# B&R Automation Studio project 67
Automation Studio 4.12.10.39

## Configuration Config1

CPU 4PP065.0571-P74, AutomationRuntime D4.52, Build 4.1.2, Vc V4.52.0

### Task classes (Cpu.sw)
```
Cyclic#1:
  Program <- Program.prg
Libraries: Library
```

### Hardware
```
4PP065_0571_P74 : 4PP065.0571-P74 v1.2.0.0
  Connector IF4:
    DNAConfiguration = manual
  Connector IF5:
    ActivateDevice = 1
  ConfigurationID = 67_Config1
  Simulation = 1
  SystemTick = 10000
  TaskClassIdleTime = 10000
```

- Physical/Config1/4PP065_0571_P74/IoMap.iom: same as Physical/Config1/4PP065_0571_P74/Cpu.per
- Physical/Config1/4PP065_0571_P74/PvMap.vvm: same as Physical/Config1/4PP065_0571_P74/Cpu.per
## Logical view

Binary libraries used (declarations not repeated): operator, runtime, astime, AsIecCon


### Program Logical/Program (ANSIC)

#### main.c - Cyclic code
```c
#include <bur/plctypes.h>

#ifdef _DEFAULT_INCLUDES
	#include <AsDefault.h>
#endif

void _CYCLIC ProgramCyclic(void)
{
	counter++;
	if (counter >= 1100)
	{
		counter = 0;
	}

	if ((counter >= 100)&&(counter < 600))
	{
		Speed = 100.0;
	}
	else
	{
		Speed = 0.0;
	}

	if (Enable)
	{
		fb_controller.e = Speed - fb_motor.w;
		FB_Regulator(&fb_controller);

		fb_motor.u = fb_controller.u;
		FB_Motor(&fb_motor);

		fb_motor2.u = Speed * fb_motor2.ke;
		FB_Motor(&fb_motor2);
	}
}
```

#### Init.c - Initialization code
```c
#include <bur/plctypes.h>

#ifdef _DEFAULT_INCLUDES
	#include <AsDefault.h>
#endif

void _INIT ProgramInit(void)
{
	//LEGO NXT

	fb_motor.tm = 0.081;
	fb_motor.ke = 0.0641;
	fb_motor.dt = 0.01;

	fb_motor.w = 0.0;
	fb_motor.phi = 0.0;
	fb_motor.integrator.in = 0.0;
	fb_motor.integrator.out = 0.0;
	fb_motor.integrator.dt = 0.01;

	fb_motor2.tm = 0.081;
	fb_motor2.ke = 0.0641;
	fb_motor2.dt = 0.01;

	fb_motor2.w = 0.0;
	fb_motor2.phi = 0.0;
	fb_motor2.integrator.in = 0.0;
	fb_motor2.integrator.out = 0.0;
	fb_motor2.integrator.dt = 0.01;

	fb_controller.k_p = 0.0052;	/* ke*Tm/Tj, Tj = 1 s */
	fb_controller.k_i = 0.0641;	/* ke/Tj */
	fb_controller.max_abs_value = 9.0;
	fb_controller.dt = 0.01;

	fb_controller.iyOld = 0.0;
	fb_controller.integrator.in = 0.0;
	fb_controller.integrator.out = 0.0;
	fb_controller.integrator.dt = 0.01;

	Speed = 0.0;
	Enable = 1;
	counter = 0;

}
```

#### Exit.c - Exit code
```c
#include <bur/plctypes.h>

#ifdef _DEFAULT_INCLUDES
	#include <AsDefault.h>
#endif

void _EXIT ProgramExit(void)
{

}
```

#### Variables.var - Local variables
```iecst
VAR
	fb_controller : {REDUND_UNREPLICABLE} FB_Regulator;
	fb_motor : {REDUND_UNREPLICABLE} FB_Motor;
	Speed : {REDUND_UNREPLICABLE} REAL;
	Enable : {REDUND_UNREPLICABLE} BOOL;
	fb_motor2 : {REDUND_UNREPLICABLE} FB_Motor;
	counter : {REDUND_UNREPLICABLE} UDINT;
END_VAR
```

### Library Logical/Library (ANSIC)

#### Library.fun - Exported functions and function blocks
```iecst
{REDUND_ERROR} {REDUND_UNREPLICABLE} FUNCTION_BLOCK FB_Integrator (*Интегратор*) (*$GROUP=User,$CAT=User,$GROUPICON=User.png,$CATICON=User.png*)
	VAR_INPUT
		in : {REDUND_UNREPLICABLE} REAL; (*Вход интегратора*)
	END_VAR
	VAR_OUTPUT
		out : {REDUND_UNREPLICABLE} REAL; (*Выход интегратора*)
	END_VAR
	VAR
		dt : {REDUND_UNREPLICABLE} REAL; (*Шаг расчёта, с*)
	END_VAR
END_FUNCTION_BLOCK

{REDUND_ERROR} {REDUND_UNREPLICABLE} FUNCTION_BLOCK FB_Motor (*Модель ДПТ*) (*$GROUP=User,$CAT=User,$GROUPICON=User.png,$CATICON=User.png*)
	VAR_INPUT
		u : {REDUND_UNREPLICABLE} REAL; (*Напряжение, В*)
	END_VAR
	VAR_OUTPUT
		w : {REDUND_UNREPLICABLE} REAL; (*Частота вращения, об/мин*)
		phi : {REDUND_UNREPLICABLE} REAL; (*Положение вала*)
	END_VAR
	VAR
		integrator : {REDUND_UNREPLICABLE} FB_Integrator; (*Интегратор*)
		tm : {REDUND_UNREPLICABLE} REAL; (*Электромеханическая постоянная времени, с*)
		ke : {REDUND_UNREPLICABLE} REAL; (*Постоянная ЭДС, В*мин/об*)
		dt : {REDUND_UNREPLICABLE} REAL; (*Шаг расчёта, с*)
	END_VAR
END_FUNCTION_BLOCK

{REDUND_ERROR} {REDUND_UNREPLICABLE} FUNCTION_BLOCK FB_Regulator (*ПИ-регулятор*) (*$GROUP=User,$CAT=User,$GROUPICON=User.png,$CATICON=User.png*)
	VAR_INPUT
		e : {REDUND_UNREPLICABLE} REAL; (*Ошибка, об/мин*)
	END_VAR
	VAR_OUTPUT
		u : {REDUND_UNREPLICABLE} REAL; (*Напряжение на ДПТ, В*)
	END_VAR
	VAR
		k_p : {REDUND_UNREPLICABLE} REAL; (*Пропорциональный коэффициент*)
		k_i : {REDUND_UNREPLICABLE} REAL; (*Интегральный коэффициент*)
		integrator : {REDUND_UNREPLICABLE} FB_Integrator; (*Интегратор*)
		iyOld : {REDUND_UNREPLICABLE} REAL; (*Интегральная составляющая*)
		max_abs_value : {REDUND_UNREPLICABLE} REAL; (*Граница ограничения, В*)
		dt : {REDUND_UNREPLICABLE} REAL; (*Шаг расчёта, с*)
	END_VAR
END_FUNCTION_BLOCK
```

#### FB_Motor.c
```c
#include <bur/plctypes.h>
#ifdef __cplusplus
	extern "C"
	{
#endif
	#include "Library.h"
#ifdef __cplusplus
	};
#endif
/* DC motor model: W(s) = 1/(ke*(Tm*s+1)) */
void FB_Motor(struct FB_Motor* inst)
{
	inst->integrator.in = (inst->u / inst->ke -  inst->w) / inst->tm;

	FB_Integrator(&inst->integrator);

	inst->w=inst->integrator.out;

	inst->phi=inst->phi + inst->w* inst->dt;
}
```

#### FB_Regulator.c
```c
#include <bur/plctypes.h>
#ifdef __cplusplus
	extern "C"
	{
#endif
	#include "Library.h"
#ifdef __cplusplus
	};
#endif
/* PI controller with output limit and anti-windup */
void FB_Regulator(struct FB_Regulator* inst)
{
	float yp;
	float y;

	yp = inst->k_p * inst->e;

	if (yp > inst->max_abs_value)
	{
		yp = inst->max_abs_value;
	}
	else if (yp < -inst->max_abs_value)
	{
		yp = -inst->max_abs_value;
	}

	y = yp+inst->iyOld;

	if (y>inst->max_abs_value)
	{
		inst->u=inst->max_abs_value;
	}
	else if (y<-inst->max_abs_value)
	{
		inst->u = -inst->max_abs_value;
	}
	else
	{
		inst->u=y;
	}

	inst->integrator.in = inst->k_i * inst->e + (inst->u - y) / inst->dt;
	inst->integrator.dt = inst->dt;
	FB_Integrator(&inst->integrator);

	inst->iyOld = inst->integrator.out;
}
```

#### FB_Integrator.c
```c
#include <bur/plctypes.h>
#ifdef __cplusplus
	extern "C"
	{
#endif
	#include "Library.h"
#ifdef __cplusplus
	};
#endif
/* Discrete integrator: out = out + in*dt */
void FB_Integrator(struct FB_Integrator* inst)
{
	inst->out = inst->out + inst->in * inst->dt;
}
```
